# EPICS StreamDevice protocol: emulation/devtest/example/example.proto
# example.proto - protocol of the fake device (fake_device.py)
Terminator = LF;

get_value { out "VAL?"; in "%f"; }
set_value { out "SET %f"; in "OK"; }
